// TIA Portal V21 export
// export: Created 2026-11-11T00:47:31.6241702Z, ExportSetting WithDefaults, DisplayName Totally Integrated Automation Portal, DisplayVersion V21 Update 3, DisplayName STEP 7 Professional, DisplayVersion V21 Update 3, DisplayName STEP 7 Safety, DisplayVersion V21, DisplayName Tech WebApplication, DisplayVersion V21, DisplayName WinCC Basic/Comfort/Advanced, DisplayVersion V21 Update 3, DisplayName WinCC Unified, DisplayVersion V21 Update 3
FUNCTION_BLOCK "FB_Fbd_ex121"   // FB132, FBD
{ S7_Optimized_Access := 'TRUE' }
VERSION : 0.1
// stored: AutoNumber true, IsIECCheckEnabled false, IsRetainMemResEnabled false, MemoryReserve 100, SetENOAutomatically false, UDAEnableTagReadback false
   VAR_INPUT
      v_mode : UInt;
      v_textid : UInt;
      v_textlistid : UInt;
   END_VAR
   VAR_OUTPUT
      v_ret_val : Int;
   END_VAR
   VAR_IN_OUT
      v_assocvalues : AssocValues;
   END_VAR
BEGIN

REGION Network 1: Gen_UsrMsg - Generate user diagnostic alarms
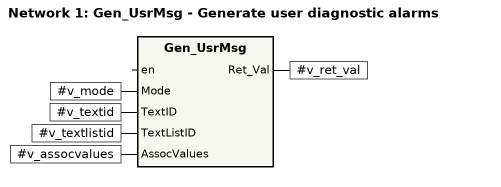
   #v_ret_val := Gen_UsrMsg(Mode := #v_mode,
                           TextID := #v_textid,
                           TextListID := #v_textlistid,
                           AssocValues := #v_assocvalues);
END_REGION
END_FUNCTION_BLOCK
